Fanuc KAREL source: kb00048.compact.KL

PROGRAM KB00048
%STACKSIZE=65535
%PRIORITY=65535
%NOLOCKGROUP
VAR
P1 : REAL
RESULT : REAL
BEGIN
P1=1.0
RESULT=COS(P1)
END KB00048
